{attribute 'linkalways'} 
{attribute 'no_explicit_call' := 'This FB is a CLASS and must be accessed using methods or properties'}
{attribute 'enable_dynamic_creation'}
FUNCTION_BLOCK _ETcWatchdogAccumulationType EXTENDS EnumDatatypeBase
VAR
	localData : ETcWatchdogAccumulationType;
	activeData : REFERENCE TO ETcWatchdogAccumulationType;
	enumBaseDatatype : _UINT(localData);
END_VAR

METHOD PRIVATE AddLocalEnumeration
VAR_INPUT
	Enumeration : T_MAXSTRING;
	Value : ETcWatchdogAccumulationType;
END_VAR
AddEnumeration(Enumeration, Value);
END_METHOD

PROPERTY PUBLIC Address : PVOID
GET
Address := ADR(activeData);
END_GET
END_PROPERTY

METHOD PUBLIC ClearReference
VAR_INPUT
END_VAR
activeData REF= localData;
SetBaseDatatypeReference();
END_METHOD

METHOD PUBLIC Clone : I_Datatype
VAR
    pClone : POINTER TO _ETcWatchdogAccumulationType;
END_VAR
pClone := __NEW(_ETcWatchdogAccumulationType(InitialValue := Value));
Clone := pClone^;
END_METHOD

METHOD FB_init : BOOL
VAR_INPUT
	bInitRetains : BOOL; // if TRUE, the retain variables are initialized (warm start / cold start)
	bInCopyCode : BOOL;  // if TRUE, the instance afterwards gets moved into the copy code (online change)
	InitialValue : ETcWatchdogAccumulationType;
END_VAR
localData := InitialValue;
AddBaseDatatype(enumBaseDatatype);
ClearReference();

AddLocalEnumeration('WD_ACC_TYPE_MEAN', ETcWatchdogAccumulationType.WD_ACC_TYPE_MEAN);
AddLocalEnumeration('WD_ACC_TYPE_PRODUCT', ETcWatchdogAccumulationType.WD_ACC_TYPE_PRODUCT);
END_METHOD

PROPERTY PUBLIC Identifier : T_MAXSTRING
GET
Identifier := 'ETcWatchdogAccumulationType';
END_GET
END_PROPERTY

METHOD IsEnumeratorValueEqual : BOOL
VAR_INPUT
	Enumerator : I_KeyValueForwardEnumerator;
END_VAR
VAR
	storedValue : ETcWatchdogAccumulationType;
END_VAR
IF NOT Enumerator.TryGet(storedValue) THEN
	RETURN;
END_IF

IsEnumeratorValueEqual := storedValue = activeData;
END_METHOD

METHOD PUBLIC MakeReferenceTo
VAR_INPUT
	ReferenceTarget : REFERENCE TO ETcWatchdogAccumulationType;
END_VAR
activeData REF= ReferenceTarget;
SetBaseDatatypeReference();
END_METHOD

METHOD PROTECTED SetBaseDatatypeReference
VAR_INPUT
END_VAR
enumBaseDatatype.MakeReferenceTo(activeData);
END_METHOD

PROPERTY PUBLIC Size : UDINT
GET
Size := SIZEOF(activeData);
END_GET
END_PROPERTY

METHOD TryMakeReferenceTo : BOOL
VAR_INPUT
	Target : I_Datatype;
END_VAR
VAR
	pTargetData : POINTER TO ETcWatchdogAccumulationType;
END_VAR
IF NOT IsEquivalentTo(Target) THEN
	RETURN;
END_IF

pTargetData := Target.Address;
activeData REF= pTargetData^;
SetBaseDatatypeReference();
TryMakeReferenceTo := TRUE;
END_METHOD

PROPERTY PUBLIC Value : ETcWatchdogAccumulationType
GET
Value := activeData;
END_GET
SET
activeData := Value;
END_SET
END_PROPERTY

END_FUNCTION_BLOCK

(* stored: Version 1.1.0.1, ProductVersion 3.1.4024.13
   POU _ETcWatchdogAccumulationType: Id {248d4af5-4761-03cb-3315-c6de778fc51d}, SpecialFunc None
   Folder Core: Id {d2b4cbb2-9a8f-0489-397b-f78d991ac3a5}
   Folder Protected: Id {16f9aa03-7ed2-03a2-0e41-96b57272633e}
   Folder Customize: Id {18c558c7-6adf-0d38-0b71-03d873f0e783}
   Folder Constructor: Id {9cf91514-1d0e-0c9f-1105-bf97c8986d40}
   Folder Private: Id {9d98cd08-4ecd-0ba2-1b23-e71709d12991}
   Folder Protected: Id {9cd420bd-0cba-0e35-1372-ae72c26a9279}
   Method AddLocalEnumeration: Id {bc0316d8-c303-020f-3200-ae372d69f243}
   Property Address: Id {c9dc5a34-c2c8-0fed-2012-7c1c7d16e6a2}
   Get Get: Id {0da831b3-b767-067c-2ed6-eba98c7a2d8e}
   Method ClearReference: Id {6ee9595e-823c-0f17-0975-11950235c338}
   Method Clone: Id {d783b119-eac7-08e7-1495-114df27e59f8}
   Method FB_init: Id {d84dcc2b-0aea-0310-3881-9d4ecee4af73}
   Property Identifier: Id {b4fd7588-94ae-05a9-0ccf-0ddee244e725}
   Get Get: Id {9d30c0f5-c52f-0a9d-395d-3bb1ee02809c}
   Method IsEnumeratorValueEqual: Id {4b28fff7-d5fa-0a61-3439-5b0d680ba79c}
   Method MakeReferenceTo: Id {d506d6b7-08c5-0f86-3479-5c7517ffa7bf}
   Method SetBaseDatatypeReference: Id {44d5e0a6-739d-0d78-2a10-48390d991e2a}
   Property Size: Id {833c6c3e-7511-0af2-33a7-ee28c6160394}
   Get Get: Id {cb49a840-9849-0bd8-3669-c894beb4bb9b}
   Method TryMakeReferenceTo: Id {a9b2d746-b49f-005d-3840-698b7489c635}
   Property Value: Id {8fa63e82-dca6-0213-0e07-7175b061756a}
   Get Get: Id {12f7bc20-aae5-0064-309b-30475507dcf4}
   Set Set: Id {37328d45-9662-00c1-18d4-b13c7c17457c} *)
